FUNCTION_BLOCK Model (* Composite Function Block Type *)
  (* Standard: 61499-2 *)
  (* Version 0.0, 7/13/2016, Andrei, nxtControl GmbH, template *)
  PACKAGE Main;
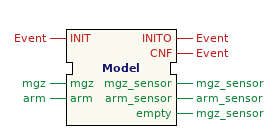
  EVENT_INPUT
    INIT; (* Initialization Request *)
  END_EVENT
  EVENT_OUTPUT
    INITO; (* Initialization Confirm *)
    CNF; (* Execution Confirmation *)
  END_EVENT
  SOCKETS
    mgz : mgz;
    arm : arm;
  END_SOCKETS
  PLUGS
    mgz_sensor : mgz_sensor;
    arm_sensor : arm_sensor;
    empty : mgz_sensor;
  END_PLUGS
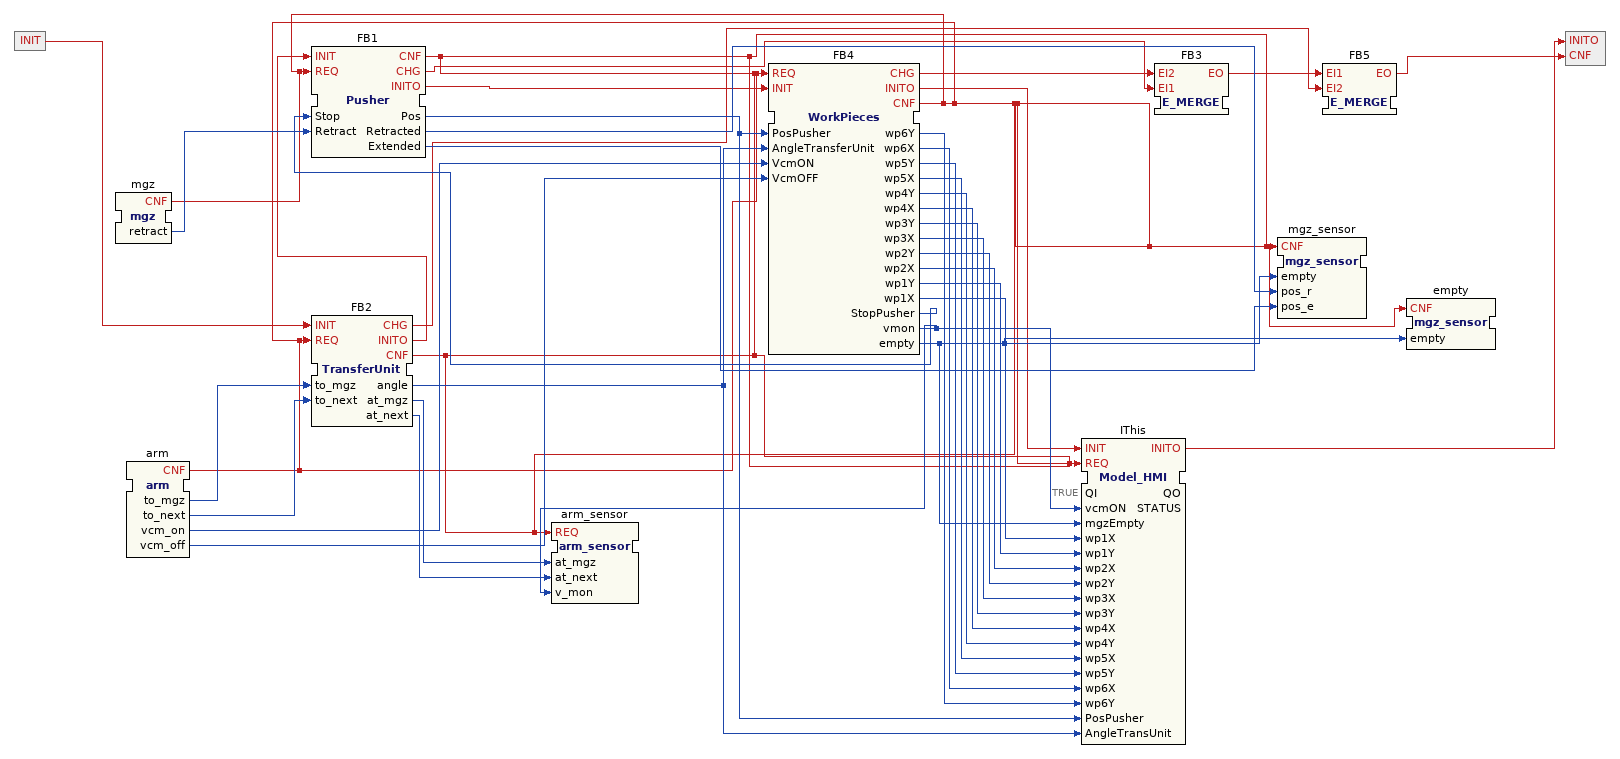
  FBS
    FB3 : E_MERGE;
    FB5 : E_MERGE;
    FB2 : TransferUnit;
    FB4 : WorkPieces;
    IThis : Model_HMI(QI := TRUE);
    FB1 : Pusher;
  END_FBS
  EVENT_CONNECTIONS
    FB1.CNF TO FB4.REQ;
    FB4.CHG TO FB3.EI2;
    FB1.CHG TO FB3.EI1;
    FB3.EO TO FB5.EI1;
    FB2.CHG TO FB5.EI2;
    FB2.INITO TO FB1.INIT;
    INIT TO FB2.INIT;
    FB1.INITO TO FB4.INIT;
    FB2.CNF TO FB4.REQ;
    FB5.EO TO CNF;
    IThis.INITO TO INITO;
    FB4.INITO TO IThis.INIT;
    FB4.CNF TO IThis.REQ;
    FB2.CNF TO IThis.REQ;
    FB1.CNF TO IThis.REQ;
    FB4.CNF TO FB1.REQ;
    FB4.CNF TO FB2.REQ;
    FB4.CNF TO mgz_sensor.CNF;
    FB1.CNF TO mgz_sensor.CNF;
    mgz.CNF TO FB1.REQ;
    arm.CNF TO FB2.REQ;
    arm.CNF TO FB4.REQ;
    FB2.CNF TO arm_sensor.REQ;
    FB4.CNF TO arm_sensor.REQ;
    FB4.CNF TO empty.CNF;
  END_CONNECTIONS
  DATA_CONNECTIONS
    FB1.Pos TO FB4.PosPusher;
    FB2.angle TO FB4.AngleTransferUnit;
    FB2.angle TO IThis.AngleTransUnit;
    FB1.Pos TO IThis.PosPusher;
    FB4.wp6Y TO IThis.wp6Y;
    FB4.wp6X TO IThis.wp6X;
    FB4.wp5Y TO IThis.wp5Y;
    FB4.wp5X TO IThis.wp5X;
    FB4.wp4Y TO IThis.wp4Y;
    FB4.wp4X TO IThis.wp4X;
    FB4.wp3Y TO IThis.wp3Y;
    FB4.wp3X TO IThis.wp3X;
    FB4.wp2Y TO IThis.wp2Y;
    FB4.wp2X TO IThis.wp2X;
    FB4.wp1Y TO IThis.wp1Y;
    FB4.wp1X TO IThis.wp1X;
    FB4.StopPusher TO FB1.Stop;
    FB4.vmon TO IThis.vcmON;
    FB4.empty TO IThis.mgzEmpty;
    FB4.empty TO mgz_sensor.empty;
    FB1.Retracted TO mgz_sensor.pos_r;
    FB1.Extended TO mgz_sensor.pos_e;
    mgz.retract TO FB1.Retract;
    arm.to_mgz TO FB2.to_mgz;
    arm.to_next TO FB2.to_next;
    arm.vcm_on TO FB4.VcmON;
    arm.vcm_off TO FB4.VcmOFF;
    FB2.at_mgz TO arm_sensor.at_mgz;
    FB2.at_next TO arm_sensor.at_next;
    FB4.vmon TO arm_sensor.v_mon;
    FB4.empty TO empty.empty;
  END_CONNECTIONS
END_FUNCTION_BLOCK
